(* IEC 61131-3 sources: plcassist-cli/packages/volt-lsp-iec/test-corpus/pro2193/Device/Plc Logic/Application/09 Misc/Library Manager/CBML, 58 files *)

(* ---- IABORTABLE.itf ---- *)
INTERFACE IABORTABLE
END_INTERFACE

(* ---- IACTIONCONTROLLER.itf ---- *)
INTERFACE IACTIONCONTROLLER
END_INTERFACE

METHOD CONTROLCLEANUPACTION
VAR_INPUT
	ITFCLEANUPACTIONPROVIDER : ICleanupActionProvider;
	XABORTPROPOSED : BOOL;
	IERRORIDPROPOSED : INT;
END_VAR
VAR_OUTPUT
	XCOMPLETE : BOOL;
	XABORT : BOOL;
	IERRORID : INT;
END_VAR
END_METHOD

METHOD CONTROLCYCLICACTION
VAR_INPUT
	ITFCYCLICACTIONPROVIDER : ICyclicActionProvider;
	ITFTIMINGCONTROLLER : ITimingController;
END_VAR
VAR_OUTPUT
	XCOMPLETE : BOOL;
	IERRORID : INT;
END_VAR
END_METHOD

METHOD CONTROLEXITACTION
VAR_INPUT
	ITFEXITACTIONPROVIDER : IExitActionProvider;
	XAFTERCLEANUP : BOOL;
	XINCOPYCODE : BOOL;
END_VAR
END_METHOD

METHOD CONTROLRESETACTION
VAR_INPUT
	ITFRESETACTIONPROVIDER : IResetActionProvider;
END_VAR
VAR_OUTPUT
	XCOMPLETE : BOOL;
END_VAR
END_METHOD

METHOD CONTROLSTARTACTION
VAR_INPUT
	ITFSTARTACTIONPROVIDER : IStartActionProvider;
END_VAR
VAR_OUTPUT
	XCOMPLETE : BOOL;
	IERRORID : INT;
END_VAR
END_METHOD

(* ---- IACTIONCONTROLLER2.itf ---- *)
INTERFACE IACTIONCONTROLLER2
END_INTERFACE

METHOD CONTROLSAMPLEACTION
VAR_INPUT
	ITFSAMPLEACTIONPROVIDER : ISampleActionProvider;
END_VAR
VAR_OUTPUT
	IERRORID : INT;
END_VAR
END_METHOD

(* ---- IACTIONPROVIDER.itf ---- *)
INTERFACE IACTIONPROVIDER
END_INTERFACE

(* ---- IBEHAVIOURMODEL.itf ---- *)
INTERFACE IBEHAVIOURMODEL
END_INTERFACE

METHOD ABORTMODEL : ERROR
VAR_INPUT
	XCOMMIT : BOOL;
END_VAR
END_METHOD

METHOD GETMODELSTATE
VAR_INPUT
	XCOMMIT : BOOL;
END_VAR
VAR_OUTPUT
	XDONE : BOOL;
	XBUSY : BOOL;
	XERROR : BOOL;
	XABORTED : BOOL;
	IERRORID : INT;
	ESTATE : STATE;
END_VAR
END_METHOD

METHOD RESETMODEL : ERROR
VAR_INPUT
	XCOMMIT : BOOL;
END_VAR
END_METHOD

METHOD STARTMODEL : ERROR
VAR_INPUT
	XCOMMIT : BOOL;
END_VAR
END_METHOD

(* ---- ICLEANUPACTIONPROVIDER.itf ---- *)
INTERFACE ICLEANUPACTIONPROVIDER
END_INTERFACE

METHOD CLEANUPACTION
VAR_INPUT
	XABORTPROPOSED : BOOL;
	IERRORIDPROPOSED : INT;
END_VAR
VAR_OUTPUT
	XCOMPLETE : BOOL;
	XABORT : BOOL;
	IERRORID : INT;
END_VAR
END_METHOD

(* ---- ICONFIGURATIONPROVIDER.itf ---- *)
INTERFACE ICONFIGURATIONPROVIDER
END_INTERFACE

METHOD GETCONFIGURATION
VAR_OUTPUT
	XLEVELCONTROLLED : BOOL;
	XTIMINGCONTROLLED : BOOL;
	XTIMELIMITED : BOOL;
	XTIMEOUTCONSTRAINT : BOOL;
	XABORTABLE : BOOL;
	XEDGETRIGGERED : BOOL;
	XHASCONTINUOUSBEHAVIOUR : BOOL;
	XSUPPORTSEXITACTION : BOOL;
END_VAR
END_METHOD

(* ---- ICONFIGURATIONPROVIDER2.itf ---- *)
INTERFACE ICONFIGURATIONPROVIDER2
END_INTERFACE

METHOD GETCONFIGURATION2
VAR_OUTPUT
	XLEVELCONTROLLED : BOOL;
	XTIMINGCONTROLLED : BOOL;
	XTIMELIMITED : BOOL;
	XTIMEOUTCONSTRAINT : BOOL;
	XABORTABLE : BOOL;
	XEDGETRIGGERED : BOOL;
	XHASCONTINUOUSBEHAVIOUR : BOOL;
	XSUPPORTSEXITACTION : BOOL;
	XSUPPORTSSAMPLEACTION : BOOL;
END_VAR
END_METHOD

(* ---- ICYCLICACTIONPROVIDER.itf ---- *)
INTERFACE ICYCLICACTIONPROVIDER
END_INTERFACE

METHOD CYCLICACTION
VAR_INPUT
	ITFTIMINGCONTROLLER : ITimingController;
END_VAR
VAR_OUTPUT
	XCOMPLETE : BOOL;
	IERRORID : INT;
END_VAR
END_METHOD

(* ---- IEDGETRIGGERED.itf ---- *)
INTERFACE IEDGETRIGGERED
END_INTERFACE

(* ---- IETRIG.itf ---- *)
INTERFACE IETRIG
END_INTERFACE

(* ---- IETRIGA.itf ---- *)
INTERFACE IETRIGA
END_INTERFACE

(* ---- IETRIGATL.itf ---- *)
INTERFACE IETRIGATL
END_INTERFACE

(* ---- IETRIGATLTO.itf ---- *)
INTERFACE IETRIGATLTO
END_INTERFACE

(* ---- IETRIGATO.itf ---- *)
INTERFACE IETRIGATO
END_INTERFACE

(* ---- IETRIGTL.itf ---- *)
INTERFACE IETRIGTL
END_INTERFACE

(* ---- IETRIGTLTO.itf ---- *)
INTERFACE IETRIGTLTO
END_INTERFACE

(* ---- IETRIGTO.itf ---- *)
INTERFACE IETRIGTO
END_INTERFACE

(* ---- IEXITACTIONPROVIDER.itf ---- *)
INTERFACE IEXITACTIONPROVIDER
END_INTERFACE

METHOD EXITACTION
VAR_INPUT
	XAFTERCLEANUP : BOOL;
	XINCOPYCODE : BOOL;
END_VAR
END_METHOD

(* ---- IHASCONTINUOUSBEHAVIOUR.itf ---- *)
INTERFACE IHASCONTINUOUSBEHAVIOUR
END_INTERFACE

(* ---- ILCON.itf ---- *)
INTERFACE ILCON
END_INTERFACE

(* ---- ILCONC.itf ---- *)
INTERFACE ILCONC
END_INTERFACE

(* ---- ILCONTL.itf ---- *)
INTERFACE ILCONTL
END_INTERFACE

(* ---- ILCONTLC.itf ---- *)
INTERFACE ILCONTLC
END_INTERFACE

(* ---- ILCONTLTO.itf ---- *)
INTERFACE ILCONTLTO
END_INTERFACE

(* ---- ILCONTO.itf ---- *)
INTERFACE ILCONTO
END_INTERFACE

(* ---- ILEVELCONTROLLED.itf ---- *)
INTERFACE ILEVELCONTROLLED
END_INTERFACE

(* ---- IRESETACTIONPROVIDER.itf ---- *)
INTERFACE IRESETACTIONPROVIDER
END_INTERFACE

METHOD RESETACTION
VAR_OUTPUT
	XCOMPLETE : BOOL;
END_VAR
END_METHOD

(* ---- ISAMPLEACTIONPROVIDER.itf ---- *)
INTERFACE ISAMPLEACTIONPROVIDER
END_INTERFACE

METHOD SAMPLEACTION
VAR_OUTPUT
	IERRORID : INT;
END_VAR
END_METHOD

(* ---- ISTARTACTIONPROVIDER.itf ---- *)
INTERFACE ISTARTACTIONPROVIDER
END_INTERFACE

METHOD STARTACTION
VAR_OUTPUT
	XCOMPLETE : BOOL;
	IERRORID : INT;
END_VAR
END_METHOD

(* ---- ITIMELIMITED.itf ---- *)
INTERFACE ITIMELIMITED
END_INTERFACE

(* ---- ITIMEOUTCONSTRAINT.itf ---- *)
INTERFACE ITIMEOUTCONSTRAINT
END_INTERFACE

(* ---- ITIMINGCONTROLLED.itf ---- *)
INTERFACE ITIMINGCONTROLLED
END_INTERFACE

(* ---- ITIMINGCONTROLLER.itf ---- *)
INTERFACE ITIMINGCONTROLLER
END_INTERFACE

METHOD CONTROLLERCHECKTIMING
VAR_OUTPUT
	XTIMEOUT : BOOL;
	XTIMELIMIT : BOOL;
END_VAR
END_METHOD

METHOD STARTINVOCATIONTIMER
END_METHOD

METHOD STARTOPERATIONTIMER
END_METHOD

(* ---- GETLIBVERSION.fun ---- *)
FUNCTION GETLIBVERSION : VERSION
END_FUNCTION

(* ---- GETLIBVERSIONNUMBER.fun ---- *)
FUNCTION GETLIBVERSIONNUMBER : DWORD
END_FUNCTION

(* ---- ISLIBRELEASED.fun ---- *)
FUNCTION ISLIBRELEASED : BOOL
END_FUNCTION

(* ---- ACTIONCONTROLLER.fb ---- *)
FUNCTION_BLOCK ACTIONCONTROLLER
END_FUNCTION_BLOCK

METHOD CONTROLCLEANUPACTION
VAR_INPUT
	ITFCLEANUPACTIONPROVIDER : ICleanupActionProvider;
	XABORTPROPOSED : BOOL;
	IERRORIDPROPOSED : INT;
END_VAR
VAR_OUTPUT
	XCOMPLETE : BOOL;
	XABORT : BOOL;
	IERRORID : INT;
END_VAR
END_METHOD

METHOD CONTROLCYCLICACTION
VAR_INPUT
	ITFCYCLICACTIONPROVIDER : ICyclicActionProvider;
	ITFTIMINGCONTROLLER : ITimingController;
END_VAR
VAR_OUTPUT
	XCOMPLETE : BOOL;
	IERRORID : INT;
END_VAR
END_METHOD

METHOD CONTROLEXITACTION
VAR_INPUT
	ITFEXITACTIONPROVIDER : IExitActionProvider;
	XAFTERCLEANUP : BOOL;
	XINCOPYCODE : BOOL;
END_VAR
END_METHOD

METHOD CONTROLRESETACTION
VAR_INPUT
	ITFRESETACTIONPROVIDER : IResetActionProvider;
END_VAR
VAR_OUTPUT
	XCOMPLETE : BOOL;
END_VAR
END_METHOD

METHOD CONTROLSAMPLEACTION
VAR_INPUT
	ITFSAMPLEACTIONPROVIDER : ISampleActionProvider;
END_VAR
VAR_OUTPUT
	IERRORID : INT;
END_VAR
END_METHOD

METHOD CONTROLSTARTACTION
VAR_INPUT
	ITFSTARTACTIONPROVIDER : IStartActionProvider;
END_VAR
VAR_OUTPUT
	XCOMPLETE : BOOL;
	IERRORID : INT;
END_VAR
END_METHOD

(* ---- BEHAVIOURMODEL.fb ---- *)
FUNCTION_BLOCK BEHAVIOURMODEL
VAR_INPUT
	ITFACTIONPROVIDER : IActionProvider;
	ITFTIMINGCONTROLLER : ITimingController;
	XCONTROL : BOOL;
	XABORT : BOOL;
	UDITIMELIMIT : UDINT;
	UDITIMEOUT : UDINT;
END_VAR
VAR_OUTPUT
	XDONE : BOOL;
	XBUSY : BOOL;
	XERROR : BOOL;
	XABORTED : BOOL;
	IERRORID : INT;
	ESTATE : STATE;
	EINTERNALERRORID : ERROR;
END_VAR
VAR
	_ITFACTIONPROVIDER : IActionProvider;
	_ITFACTIONCONTROLLER : IActionController;
	_XLEVELCONTROLLED : BOOL;
	_XTIMINGCONTROLLED : BOOL;
	_XTIMELIMITED : BOOL;
	_XTIMEOUTCONSTRAINT : BOOL;
	_XABORTABLE : BOOL;
	_XEDGETRIGGERED : BOOL;
	_XHASCONTINUOUSBEHAVIOUR : BOOL;
	_XSUPPORTSEXITACTION : BOOL;
	_XSUPPORTSSAMPLEACTION : BOOL;
	_XRESETREQUEST : BOOL;
	_XABORTPROPOSED : BOOL;
	_IERRORIDPROPOSED : INT;
	_XFIRSTHANDLESTARTINGSTATECALL : BOOL;
	_XLASTAGAIN : BOOL;
	_ITFACTIONCONTROLLER2 : IActionController2;
	_ITFSAMPLEACTIONPROVIDER : ISampleActionProvider;
	_ITFSTARTACTIONPROVIDER : IStartActionProvider;
	_ITFCYCLICACTIONPROVIDER : ICyclicActionProvider;
	_ITFCLEANUPACTIONPROVIDER : ICleanupActionProvider;
	_ITFEXITACTIONPROVIDER : IExitActionProvider;
	_ITFRESETACTIONPROVIDER : IResetActionProvider;
	ACTIONCONTROLLER : IActionController;
	MODELTIMELIMIT : UDINT;
	MODELTIMEOUT : UDINT;
END_VAR
END_FUNCTION_BLOCK

METHOD _CHECKABORTCONDITION : BOOL
END_METHOD

METHOD _CHECKPARAMETER
VAR_OUTPUT
	EERRORID : ERROR;
END_VAR
END_METHOD

METHOD _CHECKTIMEOUTCONDITION
END_METHOD

METHOD _EXECUTE
VAR_OUTPUT
	EERRORID : ERROR := ERROR.NO_ERROR;
END_VAR
END_METHOD

METHOD _RESETACTION
END_METHOD

METHOD ABORTMODEL : ERROR
VAR_INPUT
	XCOMMIT : BOOL;
END_VAR
END_METHOD

METHOD GETCONFIGURATION
VAR_OUTPUT
	XLEVELCONTROLLED : BOOL;
	XTIMINGCONTROLLED : BOOL;
	XTIMELIMITED : BOOL;
	XTIMEOUTCONSTRAINT : BOOL;
	XABORTABLE : BOOL;
	XEDGETRIGGERED : BOOL;
	XHASCONTINUOUSBEHAVIOUR : BOOL;
	XSUPPORTSEXITACTION : BOOL;
END_VAR
END_METHOD

METHOD GETCONFIGURATION2
VAR_OUTPUT
	XLEVELCONTROLLED : BOOL;
	XTIMINGCONTROLLED : BOOL;
	XTIMELIMITED : BOOL;
	XTIMEOUTCONSTRAINT : BOOL;
	XABORTABLE : BOOL;
	XEDGETRIGGERED : BOOL;
	XHASCONTINUOUSBEHAVIOUR : BOOL;
	XSUPPORTSEXITACTION : BOOL;
	XSUPPORTSSAMPLEACTION : BOOL;
END_VAR
END_METHOD

METHOD GETMODELSTATE
VAR_INPUT
	XCOMMIT : BOOL;
END_VAR
VAR_OUTPUT
	XDONE : BOOL;
	XBUSY : BOOL;
	XERROR : BOOL;
	XABORTED : BOOL;
	IERRORID : INT;
	ESTATE : STATE;
END_VAR
END_METHOD

METHOD RESETMODEL : ERROR
VAR_INPUT
	XCOMMIT : BOOL;
END_VAR
END_METHOD

METHOD STARTMODEL : ERROR
VAR_INPUT
	XCOMMIT : BOOL;
END_VAR
END_METHOD

METHOD _HANDLEABORTEDSTATE
VAR_OUTPUT
	XAGAIN : BOOL;
END_VAR
END_METHOD

METHOD _HANDLECLEANINGSTATE
VAR_OUTPUT
	XAGAIN : BOOL;
END_VAR
END_METHOD

METHOD _HANDLEDONESTATE
VAR_OUTPUT
	XAGAIN : BOOL;
END_VAR
END_METHOD

METHOD _HANDLEDORMANTSTATE
VAR_OUTPUT
	XAGAIN : BOOL;
END_VAR
END_METHOD

METHOD _HANDLEERRORSTATE
VAR_OUTPUT
	XAGAIN : BOOL;
END_VAR
END_METHOD

METHOD _HANDLEEXECUTINGSTATE
VAR_OUTPUT
	XAGAIN : BOOL;
END_VAR
END_METHOD

METHOD _HANDLERESETTINGSTATE
VAR_OUTPUT
	XAGAIN : BOOL;
END_VAR
END_METHOD

METHOD _HANDLESTARTINGSTATE
VAR_OUTPUT
	XAGAIN : BOOL;
	IERRORID : INT;
END_VAR
END_METHOD

METHOD _STATEMACHINE : ERROR
END_METHOD

(* ---- BEHAVIOURMODELBASE.fb ---- *)
FUNCTION_BLOCK BEHAVIOURMODELBASE
VAR
	_MODEL : BehaviourModel := STRUCT(itfActionProvider := THIS^, itfTimingController := 0);
	ACTIONCONTROLLER : IActionController;
	MODELTIMELIMIT : UDINT;
	MODELTIMEOUT : UDINT;
END_VAR
END_FUNCTION_BLOCK

METHOD FB_EXIT : BOOL
VAR_INPUT
	BINCOPYCODE : BOOL;
END_VAR
END_METHOD

METHOD _EXECUTE
VAR_OUTPUT
	EERRORID : ERROR;
END_VAR
END_METHOD

METHOD CLEANUPACTION
VAR_INPUT
	XABORTPROPOSED : BOOL;
	IERRORIDPROPOSED : INT;
END_VAR
VAR_OUTPUT
	XCOMPLETE : BOOL := TRUE;
	XABORT : BOOL := xAbortProposed;
	IERRORID : INT := iErrorIDProposed;
END_VAR
END_METHOD

METHOD CYCLICACTION
VAR_INPUT
	ITFTIMINGCONTROLLER : ITimingController;
END_VAR
VAR_OUTPUT
	XCOMPLETE : BOOL := TRUE;
	IERRORID : INT := 0;
END_VAR
END_METHOD

METHOD EXITACTION
VAR_INPUT
	XAFTERCLEANUP : BOOL;
	XINCOPYCODE : BOOL;
END_VAR
END_METHOD

METHOD RESETACTION
VAR_OUTPUT
	XCOMPLETE : BOOL := TRUE;
END_VAR
END_METHOD

METHOD STARTACTION
VAR_OUTPUT
	XCOMPLETE : BOOL := TRUE;
	IERRORID : INT := 0;
END_VAR
END_METHOD

METHOD ABORTMODEL : ERROR
VAR_INPUT
	XCOMMIT : BOOL;
END_VAR
END_METHOD

METHOD GETCONFIGURATION
VAR_OUTPUT
	XLEVELCONTROLLED : BOOL;
	XTIMINGCONTROLLED : BOOL;
	XTIMELIMITED : BOOL;
	XTIMEOUTCONSTRAINT : BOOL;
	XABORTABLE : BOOL;
	XEDGETRIGGERED : BOOL;
	XHASCONTINUOUSBEHAVIOUR : BOOL;
	XSUPPORTSEXITACTION : BOOL;
END_VAR
END_METHOD

METHOD GETCONFIGURATION2
VAR_OUTPUT
	XLEVELCONTROLLED : BOOL;
	XTIMINGCONTROLLED : BOOL;
	XTIMELIMITED : BOOL;
	XTIMEOUTCONSTRAINT : BOOL;
	XABORTABLE : BOOL;
	XEDGETRIGGERED : BOOL;
	XHASCONTINUOUSBEHAVIOUR : BOOL;
	XSUPPORTSEXITACTION : BOOL;
	XSUPPORTSSAMPLEACTION : BOOL;
END_VAR
END_METHOD

METHOD GETMODELSTATE
VAR_INPUT
	XCOMMIT : BOOL;
END_VAR
VAR_OUTPUT
	XDONE : BOOL;
	XBUSY : BOOL;
	XERROR : BOOL;
	XABORTED : BOOL;
	IERRORID : INT;
	ESTATE : STATE;
END_VAR
END_METHOD

METHOD RESETMODEL : ERROR
VAR_INPUT
	XCOMMIT : BOOL;
END_VAR
END_METHOD

METHOD STARTMODEL : ERROR
VAR_INPUT
	XCOMMIT : BOOL;
END_VAR
END_METHOD

(* ---- EDGETRIGGEREDBEHAVIOURMODELBASE.fb ---- *)
FUNCTION_BLOCK EDGETRIGGEREDBEHAVIOURMODELBASE EXTENDS BehaviourModelBase
END_FUNCTION_BLOCK

METHOD SAMPLEACTION
VAR_OUTPUT
	IERRORID : INT := 0;
END_VAR
END_METHOD

(* ---- EDGETRIGGEREDTIMINGCONTROLLEDBEHAVIOURMODELBASE.fb ---- *)
FUNCTION_BLOCK EDGETRIGGEREDTIMINGCONTROLLEDBEHAVIOURMODELBASE EXTENDS TimingControlledBehaviourModelBase
END_FUNCTION_BLOCK

METHOD SAMPLEACTION
VAR_OUTPUT
	IERRORID : INT := 0;
END_VAR
END_METHOD

(* ---- ETRIG.fb ---- *)
FUNCTION_BLOCK ETRIG EXTENDS EdgeTriggeredBehaviourModelBase
VAR_INPUT
	XEXECUTE : BOOL;
END_VAR
VAR_OUTPUT
	XDONE : BOOL;
	XBUSY : BOOL;
	XERROR : BOOL;
END_VAR
END_FUNCTION_BLOCK

METHOD _EXECUTE
VAR_OUTPUT
	EERRORID : ERROR;
END_VAR
END_METHOD

METHOD GETMODELSTATE
VAR_INPUT
	XCOMMIT : BOOL;
END_VAR
VAR_OUTPUT
	XDONE : BOOL;
	XBUSY : BOOL;
	XERROR : BOOL;
	XABORTED : BOOL;
	IERRORID : INT;
	ESTATE : STATE;
END_VAR
END_METHOD

METHOD RESETMODEL : ERROR
VAR_INPUT
	XCOMMIT : BOOL;
END_VAR
END_METHOD

METHOD STARTMODEL : ERROR
VAR_INPUT
	XCOMMIT : BOOL;
END_VAR
END_METHOD

(* ---- ETRIGA.fb ---- *)
FUNCTION_BLOCK ETRIGA EXTENDS ETrig
VAR_INPUT
	XABORT : BOOL;
END_VAR
VAR_OUTPUT
	XABORTED : BOOL;
END_VAR
END_FUNCTION_BLOCK

METHOD _EXECUTE
VAR_OUTPUT
	EERRORID : ERROR;
END_VAR
END_METHOD

METHOD ABORTMODEL : ERROR
VAR_INPUT
	XCOMMIT : BOOL;
END_VAR
END_METHOD

METHOD GETMODELSTATE
VAR_INPUT
	XCOMMIT : BOOL;
END_VAR
VAR_OUTPUT
	XDONE : BOOL;
	XBUSY : BOOL;
	XERROR : BOOL;
	XABORTED : BOOL;
	IERRORID : INT;
	ESTATE : STATE;
END_VAR
END_METHOD

METHOD RESETMODEL : ERROR
VAR_INPUT
	XCOMMIT : BOOL;
END_VAR
END_METHOD

(* ---- ETRIGATL.fb ---- *)
FUNCTION_BLOCK ETRIGATL EXTENDS EdgeTriggeredTimingControlledBehaviourModelBase
VAR_INPUT
	XEXECUTE : BOOL;
	XABORT : BOOL;
	UDITIMELIMIT : UDINT;
END_VAR
VAR_OUTPUT
	XDONE : BOOL;
	XBUSY : BOOL;
	XERROR : BOOL;
	XABORTED : BOOL;
END_VAR
VAR
	MODELTIMELIMIT : UDINT;
END_VAR
END_FUNCTION_BLOCK

METHOD _EXECUTE
VAR_OUTPUT
	EERRORID : ERROR;
END_VAR
END_METHOD

METHOD ABORTMODEL : ERROR
VAR_INPUT
	XCOMMIT : BOOL;
END_VAR
END_METHOD

METHOD GETMODELSTATE
VAR_INPUT
	XCOMMIT : BOOL;
END_VAR
VAR_OUTPUT
	XDONE : BOOL;
	XBUSY : BOOL;
	XERROR : BOOL;
	XABORTED : BOOL;
	IERRORID : INT;
	ESTATE : STATE;
END_VAR
END_METHOD

METHOD RESETMODEL : ERROR
VAR_INPUT
	XCOMMIT : BOOL;
END_VAR
END_METHOD

METHOD STARTMODEL : ERROR
VAR_INPUT
	XCOMMIT : BOOL;
END_VAR
END_METHOD

(* ---- ETRIGATLTO.fb ---- *)
FUNCTION_BLOCK ETRIGATLTO EXTENDS ETrigATl
VAR_INPUT
	UDITIMEOUT : UDINT;
END_VAR
VAR
	MODELTIMEOUT : UDINT;
END_VAR
END_FUNCTION_BLOCK

METHOD _EXECUTE
VAR_OUTPUT
	EERRORID : ERROR;
END_VAR
END_METHOD

METHOD GETMODELSTATE
VAR_INPUT
	XCOMMIT : BOOL;
END_VAR
VAR_OUTPUT
	XDONE : BOOL;
	XBUSY : BOOL;
	XERROR : BOOL;
	XABORTED : BOOL;
	IERRORID : INT;
	ESTATE : STATE;
END_VAR
END_METHOD

(* ---- ETRIGATO.fb ---- *)
FUNCTION_BLOCK ETRIGATO EXTENDS EdgeTriggeredTimingControlledBehaviourModelBase
VAR_INPUT
	XEXECUTE : BOOL;
	XABORT : BOOL;
	UDITIMEOUT : UDINT;
END_VAR
VAR_OUTPUT
	XDONE : BOOL;
	XBUSY : BOOL;
	XERROR : BOOL;
	XABORTED : BOOL;
END_VAR
VAR
	MODELTIMEOUT : UDINT;
END_VAR
END_FUNCTION_BLOCK

METHOD _EXECUTE
VAR_OUTPUT
	EERRORID : ERROR;
END_VAR
END_METHOD

METHOD ABORTMODEL : ERROR
VAR_INPUT
	XCOMMIT : BOOL;
END_VAR
END_METHOD

METHOD GETMODELSTATE
VAR_INPUT
	XCOMMIT : BOOL;
END_VAR
VAR_OUTPUT
	XDONE : BOOL;
	XBUSY : BOOL;
	XERROR : BOOL;
	XABORTED : BOOL;
	IERRORID : INT;
	ESTATE : STATE;
END_VAR
END_METHOD

METHOD RESETMODEL : ERROR
VAR_INPUT
	XCOMMIT : BOOL;
END_VAR
END_METHOD

METHOD STARTMODEL : ERROR
VAR_INPUT
	XCOMMIT : BOOL;
END_VAR
END_METHOD

(* ---- ETRIGTL.fb ---- *)
FUNCTION_BLOCK ETRIGTL EXTENDS EdgeTriggeredTimingControlledBehaviourModelBase
VAR_INPUT
	XEXECUTE : BOOL;
	UDITIMELIMIT : UDINT;
END_VAR
VAR_OUTPUT
	XDONE : BOOL;
	XBUSY : BOOL;
	XERROR : BOOL;
END_VAR
VAR
	MODELTIMELIMIT : UDINT;
END_VAR
END_FUNCTION_BLOCK

METHOD _EXECUTE
VAR_OUTPUT
	EERRORID : ERROR;
END_VAR
END_METHOD

METHOD GETMODELSTATE
VAR_INPUT
	XCOMMIT : BOOL;
END_VAR
VAR_OUTPUT
	XDONE : BOOL;
	XBUSY : BOOL;
	XERROR : BOOL;
	XABORTED : BOOL;
	IERRORID : INT;
	ESTATE : STATE;
END_VAR
END_METHOD

METHOD RESETMODEL : ERROR
VAR_INPUT
	XCOMMIT : BOOL;
END_VAR
END_METHOD

METHOD STARTMODEL : ERROR
VAR_INPUT
	XCOMMIT : BOOL;
END_VAR
END_METHOD

(* ---- ETRIGTLTO.fb ---- *)
FUNCTION_BLOCK ETRIGTLTO EXTENDS ETrigTl
VAR_INPUT
	UDITIMEOUT : UDINT;
END_VAR
VAR
	MODELTIMEOUT : UDINT;
END_VAR
END_FUNCTION_BLOCK

METHOD _EXECUTE
VAR_OUTPUT
	EERRORID : ERROR;
END_VAR
END_METHOD

METHOD GETMODELSTATE
VAR_INPUT
	XCOMMIT : BOOL;
END_VAR
VAR_OUTPUT
	XDONE : BOOL;
	XBUSY : BOOL;
	XERROR : BOOL;
	XABORTED : BOOL;
	IERRORID : INT;
	ESTATE : STATE;
END_VAR
END_METHOD

(* ---- ETRIGTO.fb ---- *)
FUNCTION_BLOCK ETRIGTO EXTENDS EdgeTriggeredTimingControlledBehaviourModelBase
VAR_INPUT
	XEXECUTE : BOOL;
	UDITIMEOUT : UDINT;
END_VAR
VAR_OUTPUT
	XDONE : BOOL;
	XBUSY : BOOL;
	XERROR : BOOL;
END_VAR
VAR
	MODELTIMEOUT : UDINT;
END_VAR
END_FUNCTION_BLOCK

METHOD _EXECUTE
VAR_OUTPUT
	EERRORID : ERROR;
END_VAR
END_METHOD

METHOD GETMODELSTATE
VAR_INPUT
	XCOMMIT : BOOL;
END_VAR
VAR_OUTPUT
	XDONE : BOOL;
	XBUSY : BOOL;
	XERROR : BOOL;
	XABORTED : BOOL;
	IERRORID : INT;
	ESTATE : STATE;
END_VAR
END_METHOD

METHOD RESETMODEL : ERROR
VAR_INPUT
	XCOMMIT : BOOL;
END_VAR
END_METHOD

METHOD STARTMODEL : ERROR
VAR_INPUT
	XCOMMIT : BOOL;
END_VAR
END_METHOD

(* ---- LCON.fb ---- *)
FUNCTION_BLOCK LCON EXTENDS BehaviourModelBase
VAR_INPUT
	XENABLE : BOOL;
END_VAR
VAR_OUTPUT
	XDONE : BOOL;
	XBUSY : BOOL;
	XERROR : BOOL;
END_VAR
END_FUNCTION_BLOCK

METHOD _EXECUTE
VAR_OUTPUT
	EERRORID : ERROR;
END_VAR
END_METHOD

METHOD ABORTMODEL : ERROR
VAR_INPUT
	XCOMMIT : BOOL;
END_VAR
END_METHOD

METHOD GETMODELSTATE
VAR_INPUT
	XCOMMIT : BOOL;
END_VAR
VAR_OUTPUT
	XDONE : BOOL;
	XBUSY : BOOL;
	XERROR : BOOL;
	XABORTED : BOOL;
	IERRORID : INT;
	ESTATE : STATE;
END_VAR
END_METHOD

METHOD RESETMODEL : ERROR
VAR_INPUT
	XCOMMIT : BOOL;
END_VAR
END_METHOD

METHOD STARTMODEL : ERROR
VAR_INPUT
	XCOMMIT : BOOL;
END_VAR
END_METHOD

(* ---- LCONC.fb ---- *)
FUNCTION_BLOCK LCONC EXTENDS BehaviourModelBase
VAR_INPUT
	XENABLE : BOOL;
END_VAR
VAR_OUTPUT
	XBUSY : BOOL;
	XERROR : BOOL;
END_VAR
END_FUNCTION_BLOCK

METHOD _EXECUTE
VAR_OUTPUT
	EERRORID : ERROR;
END_VAR
END_METHOD

METHOD ABORTMODEL : ERROR
VAR_INPUT
	XCOMMIT : BOOL;
END_VAR
END_METHOD

METHOD GETMODELSTATE
VAR_INPUT
	XCOMMIT : BOOL;
END_VAR
VAR_OUTPUT
	XDONE : BOOL;
	XBUSY : BOOL;
	XERROR : BOOL;
	XABORTED : BOOL;
	IERRORID : INT;
	ESTATE : STATE;
END_VAR
END_METHOD

METHOD RESETMODEL : ERROR
VAR_INPUT
	XCOMMIT : BOOL;
END_VAR
END_METHOD

METHOD STARTMODEL : ERROR
VAR_INPUT
	XCOMMIT : BOOL;
END_VAR
END_METHOD

(* ---- LCONTL.fb ---- *)
FUNCTION_BLOCK LCONTL EXTENDS TimingControlledBehaviourModelBase
VAR_INPUT
	XENABLE : BOOL;
	UDITIMELIMIT : UDINT;
END_VAR
VAR_OUTPUT
	XDONE : BOOL;
	XBUSY : BOOL;
	XERROR : BOOL;
END_VAR
VAR
	MODELTIMELIMIT : UDINT;
END_VAR
END_FUNCTION_BLOCK

METHOD _EXECUTE
VAR_OUTPUT
	EERRORID : ERROR;
END_VAR
END_METHOD

METHOD ABORTMODEL : ERROR
VAR_INPUT
	XCOMMIT : BOOL;
END_VAR
END_METHOD

METHOD GETMODELSTATE
VAR_INPUT
	XCOMMIT : BOOL;
END_VAR
VAR_OUTPUT
	XDONE : BOOL;
	XBUSY : BOOL;
	XERROR : BOOL;
	XABORTED : BOOL;
	IERRORID : INT;
	ESTATE : STATE;
END_VAR
END_METHOD

METHOD RESETMODEL : ERROR
VAR_INPUT
	XCOMMIT : BOOL;
END_VAR
END_METHOD

METHOD STARTMODEL : ERROR
VAR_INPUT
	XCOMMIT : BOOL;
END_VAR
END_METHOD

(* ---- LCONTLC.fb ---- *)
FUNCTION_BLOCK LCONTLC EXTENDS TimingControlledBehaviourModelBase
VAR_INPUT
	XENABLE : BOOL;
	UDITIMELIMIT : UDINT;
END_VAR
VAR_OUTPUT
	XBUSY : BOOL;
	XERROR : BOOL;
END_VAR
VAR
	MODELTIMELIMIT : UDINT;
END_VAR
END_FUNCTION_BLOCK

METHOD _EXECUTE
VAR_OUTPUT
	EERRORID : ERROR;
END_VAR
END_METHOD

METHOD ABORTMODEL : ERROR
VAR_INPUT
	XCOMMIT : BOOL;
END_VAR
END_METHOD

METHOD GETMODELSTATE
VAR_INPUT
	XCOMMIT : BOOL;
END_VAR
VAR_OUTPUT
	XDONE : BOOL;
	XBUSY : BOOL;
	XERROR : BOOL;
	XABORTED : BOOL;
	IERRORID : INT;
	ESTATE : STATE;
END_VAR
END_METHOD

METHOD RESETMODEL : ERROR
VAR_INPUT
	XCOMMIT : BOOL;
END_VAR
END_METHOD

METHOD STARTMODEL : ERROR
VAR_INPUT
	XCOMMIT : BOOL;
END_VAR
END_METHOD

(* ---- LCONTLTO.fb ---- *)
FUNCTION_BLOCK LCONTLTO EXTENDS LConTl
VAR_INPUT
	UDITIMEOUT : UDINT;
END_VAR
VAR
	MODELTIMEOUT : UDINT;
END_VAR
END_FUNCTION_BLOCK

METHOD _EXECUTE
VAR_OUTPUT
	EERRORID : ERROR;
END_VAR
END_METHOD

METHOD GETMODELSTATE
VAR_INPUT
	XCOMMIT : BOOL;
END_VAR
VAR_OUTPUT
	XDONE : BOOL;
	XBUSY : BOOL;
	XERROR : BOOL;
	XABORTED : BOOL;
	IERRORID : INT;
	ESTATE : STATE;
END_VAR
END_METHOD

(* ---- LCONTO.fb ---- *)
FUNCTION_BLOCK LCONTO EXTENDS TimingControlledBehaviourModelBase
VAR_INPUT
	XENABLE : BOOL;
	UDITIMEOUT : UDINT;
END_VAR
VAR_OUTPUT
	XDONE : BOOL;
	XBUSY : BOOL;
	XERROR : BOOL;
END_VAR
VAR
	MODELTIMEOUT : UDINT;
END_VAR
END_FUNCTION_BLOCK

METHOD _EXECUTE
VAR_OUTPUT
	EERRORID : ERROR;
END_VAR
END_METHOD

METHOD ABORTMODEL : ERROR
VAR_INPUT
	XCOMMIT : BOOL;
END_VAR
END_METHOD

METHOD GETMODELSTATE
VAR_INPUT
	XCOMMIT : BOOL;
END_VAR
VAR_OUTPUT
	XDONE : BOOL;
	XBUSY : BOOL;
	XERROR : BOOL;
	XABORTED : BOOL;
	IERRORID : INT;
	ESTATE : STATE;
END_VAR
END_METHOD

METHOD RESETMODEL : ERROR
VAR_INPUT
	XCOMMIT : BOOL;
END_VAR
END_METHOD

METHOD STARTMODEL : ERROR
VAR_INPUT
	XCOMMIT : BOOL;
END_VAR
END_METHOD

(* ---- TIMINGCONTROLLEDBEHAVIOURMODELBASE.fb ---- *)
FUNCTION_BLOCK TIMINGCONTROLLEDBEHAVIOURMODELBASE
VAR
	_TIMINGCONTROLLER : TimingController;
	_MODEL : BehaviourModel := STRUCT(itfActionProvider := THIS^, itfTimingController := _TimingController);
	ACTIONCONTROLLER : IActionController;
	MODELTIMELIMIT : UDINT;
	MODELTIMEOUT : UDINT;
END_VAR
END_FUNCTION_BLOCK

METHOD FB_EXIT : BOOL
VAR_INPUT
	BINCOPYCODE : BOOL;
END_VAR
END_METHOD

METHOD _EXECUTE
VAR_OUTPUT
	EERRORID : ERROR;
END_VAR
END_METHOD

METHOD CLEANUPACTION
VAR_INPUT
	XABORTPROPOSED : BOOL;
	IERRORIDPROPOSED : INT;
END_VAR
VAR_OUTPUT
	XCOMPLETE : BOOL := TRUE;
	XABORT : BOOL := xAbortProposed;
	IERRORID : INT := iErrorIDProposed;
END_VAR
END_METHOD

METHOD CYCLICACTION
VAR_INPUT
	ITFTIMINGCONTROLLER : ITimingController;
END_VAR
VAR_OUTPUT
	XCOMPLETE : BOOL := TRUE;
	IERRORID : INT := 0;
END_VAR
END_METHOD

METHOD EXITACTION
VAR_INPUT
	XAFTERCLEANUP : BOOL;
	XINCOPYCODE : BOOL;
END_VAR
END_METHOD

METHOD RESETACTION
VAR_OUTPUT
	XCOMPLETE : BOOL := TRUE;
END_VAR
END_METHOD

METHOD STARTACTION
VAR_OUTPUT
	XCOMPLETE : BOOL := TRUE;
	IERRORID : INT := 0;
END_VAR
END_METHOD

METHOD ABORTMODEL : ERROR
VAR_INPUT
	XCOMMIT : BOOL;
END_VAR
END_METHOD

METHOD GETCONFIGURATION
VAR_OUTPUT
	XLEVELCONTROLLED : BOOL;
	XTIMINGCONTROLLED : BOOL;
	XTIMELIMITED : BOOL;
	XTIMEOUTCONSTRAINT : BOOL;
	XABORTABLE : BOOL;
	XEDGETRIGGERED : BOOL;
	XHASCONTINUOUSBEHAVIOUR : BOOL;
	XSUPPORTSEXITACTION : BOOL;
END_VAR
END_METHOD

METHOD GETCONFIGURATION2
VAR_OUTPUT
	XLEVELCONTROLLED : BOOL;
	XTIMINGCONTROLLED : BOOL;
	XTIMELIMITED : BOOL;
	XTIMEOUTCONSTRAINT : BOOL;
	XABORTABLE : BOOL;
	XEDGETRIGGERED : BOOL;
	XHASCONTINUOUSBEHAVIOUR : BOOL;
	XSUPPORTSEXITACTION : BOOL;
	XSUPPORTSSAMPLEACTION : BOOL;
END_VAR
END_METHOD

METHOD GETMODELSTATE
VAR_INPUT
	XCOMMIT : BOOL;
END_VAR
VAR_OUTPUT
	XDONE : BOOL;
	XBUSY : BOOL;
	XERROR : BOOL;
	XABORTED : BOOL;
	IERRORID : INT;
	ESTATE : STATE;
END_VAR
END_METHOD

METHOD RESETMODEL : ERROR
VAR_INPUT
	XCOMMIT : BOOL;
END_VAR
END_METHOD

METHOD STARTMODEL : ERROR
VAR_INPUT
	XCOMMIT : BOOL;
END_VAR
END_METHOD

(* ---- TIMINGCONTROLLER.fb ---- *)
FUNCTION_BLOCK TIMINGCONTROLLER
VAR
	_UDITIMELIMIT : UDINT;
	_UDITIMEOUT : UDINT;
	_UDIOPERATIONSTARTTIME : UDINT;
	_UDIINVOCATIONSTARTTIME : UDINT;
	CONTROLLERTIMELIMIT : UDINT;
	CONTROLLERTIMEOUT : UDINT;
	CURRENTCONTROLLERTIME : UDINT;
END_VAR
END_FUNCTION_BLOCK

METHOD CONTROLLERCHECKTIMING
VAR_OUTPUT
	XTIMEOUT : BOOL;
	XTIMELIMIT : BOOL;
END_VAR
END_METHOD

METHOD STARTINVOCATIONTIMER
END_METHOD

METHOD STARTOPERATIONTIMER
END_METHOD
